// TIA Portal V21 export
// export: Created 2026-11-11T00:48:07.5313915Z, ExportSetting WithDefaults, DisplayName Totally Integrated Automation Portal, DisplayVersion V21 Update 3, DisplayName STEP 7 Professional, DisplayVersion V21 Update 3, DisplayName STEP 7 Safety, DisplayVersion V21, DisplayName Tech WebApplication, DisplayVersion V21, DisplayName WinCC Basic/Comfort/Advanced, DisplayVersion V21 Update 3, DisplayName WinCC Unified, DisplayVersion V21 Update 3
FUNCTION_BLOCK "FB_Scl_sl003"   // FB23, SCL
{ S7_Optimized_Access := 'TRUE' }
VERSION : 0.1
// stored: AutoNumber true, IsIECCheckEnabled false, IsRetainMemResEnabled false, MemoryReserve 100, SetENOAutomatically false, UDAEnableTagReadback false
   VAR_INPUT
      v_in : Bool;
      v_pt : Time;
   END_VAR
   VAR_OUTPUT
      v_q : Bool;
      v_et : Time;
   END_VAR
   VAR
      inst { S7_SetPoint := 'True'} : TP_TIME;
   END_VAR
BEGIN
   #inst(IN := #v_in, PT := #v_pt, Q => #v_q, ET => #v_et);
END_FUNCTION_BLOCK
